// LS Electric XG5000 project: FSS
// PLC LSPLCXBMDN16H2
// module base 0 slot 0: 입출력 모듈:XBM-DN/DP16H2 (DC 24V입력, 트랜지스터 출력 16점)
// module base 0 slot 1: 내장위치결정:XBF-PO02E (오픈컬렉터형, 2축)
// module base 0 slot 2: 아날로그출력 모듈:XBF-DC04A (D/A 전류 출력형 4채널)
// module base 0 slot 3: 아날로그출력 모듈:XBF-DC04A (D/A 전류 출력형 4채널)

PROGRAM NewProgram (task: 스캔 프로그램)

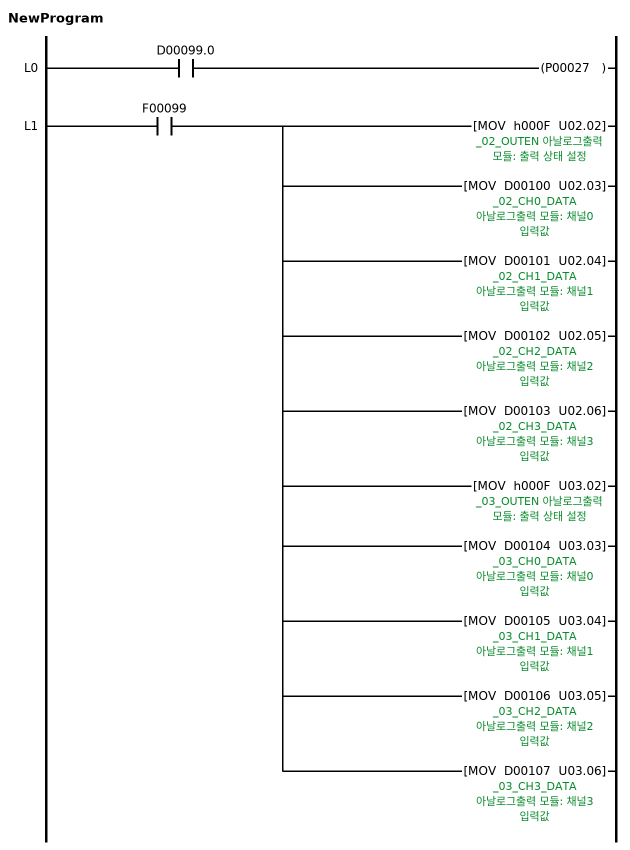
; L0
LOAD      D00099.0
OUT       P00027
; L1
LOAD      F00099
MOV       h000F U02.02	// _02_OUTEN 아날로그출력 모듈: 출력 상태 설정
MOV       D00100 U02.03	// _02_CH0_DATA 아날로그출력 모듈: 채널0 입력값
MOV       D00101 U02.04	// _02_CH1_DATA 아날로그출력 모듈: 채널1 입력값
MOV       D00102 U02.05	// _02_CH2_DATA 아날로그출력 모듈: 채널2 입력값
MOV       D00103 U02.06	// _02_CH3_DATA 아날로그출력 모듈: 채널3 입력값
MOV       h000F U03.02	// _03_OUTEN 아날로그출력 모듈: 출력 상태 설정
MOV       D00104 U03.03	// _03_CH0_DATA 아날로그출력 모듈: 채널0 입력값
MOV       D00105 U03.04	// _03_CH1_DATA 아날로그출력 모듈: 채널1 입력값
MOV       D00106 U03.05	// _03_CH2_DATA 아날로그출력 모듈: 채널2 입력값
MOV       D00107 U03.06	// _03_CH3_DATA 아날로그출력 모듈: 채널3 입력값